GLOBALCONSTANTS FuncConst (* Konstanten fuer Function-Aufruf-Uebung *)
  (* Standard: 61499-1; Description: Copyright (c) 2026 Meisterschulen am Ostbahnhof This program and the accompanying materials are made available under the terms of the Eclipse Public License 2.0 which is available at https://www.eclipse.org/legal/epl-2.0/ SPDX-License-Identifier: EPL-2.0 *)
  (* Version 1.0, 2026-10-16, Franz Höpfinger, Meisterschulen am Ostbahnhof, Uebung: Function aus GCF aufrufen *)
  PACKAGE Meins::GcfFunctionCall::const;
  VAR_GLOBAL CONSTANT
    BASE_VALUE : INT := 7;
    DOUBLE_VALUE : INT := Meins::GcfFunctionCall::F_Double(BASE_VALUE); (* Aufruf F_Double in GCF *)
  END_VAR
END_GLOBALCONSTANTS
